(* IEC 61131-3 sources: Versio-VersionControlSystem/fixtures/projects/MachineWithMembers/Device/Plc Logic/Application/Pumps/FB_Pump, 1 file *)

(* ---- Start.st ---- *)
METHOD Start : BOOL
VAR_INPUT
	target : INT;
END_VAR

// --- BEGIN IMPLEMENTATION ---

speed := target;
Start := TRUE;
